(* Communikation structure from drive to plc *)

TYPE ST_STOEBERSI6SC6CIA402TOPLC_1 :
STRUCT
	snA542ModesOfOperationDisplay		:SINT;
	dnA545PositionActualValue			:DINT;
	dnA553VelocityActualValue 			:DINT;
	nA564TorqueActualValue 				:INT;
	dw1A636DigitalInputs				:DWORD;
	dnA620AdditionalPositionActualValue	:DINT;
	wE201Statuswort2 					:WORD;
	wA67UserStatuswort 					:WORD;
END_STRUCT
END_TYPE

(* stored: Version 1.1.0.1, ProductVersion 3.1.4024.15
   DUT ST_STOEBERSI6SC6CIA402TOPLC_1: Id {f532bbf8-d4dd-492a-8356-6003871f18f4} *)
